Fanuc KAREL source: KT00511.KL

PROGRAM KT00511
%NOLOCKGROUP
VAR
  P1: XYZWPR
  P2: JOINTPOS
  OUT: XYZWPREXT
BEGIN
  P1.X = 1.0
  OUT = P1 : P2
END KT00511
